TYPE ST_LightInfo :
STRUCT
    sLocationId : STRING(16);
    {attribute 'TcEncoding' := 'UTF-8'}
    sLocationName : STRING(64);
    sId : STRING(16);
    {attribute 'TcEncoding' := 'UTF-8'}
    sName : STRING(64);
    sType : STRING(16) := 'light';
    bOn : BOOL;
END_STRUCT
END_TYPE

(* stored: Version 1.1.0.1
   DUT ST_LightInfo: Id {16c391bc-c288-45f3-aefa-07ee4b479fa7} *)
